Yaskawa INFORM job: OVERLAP3.JBI

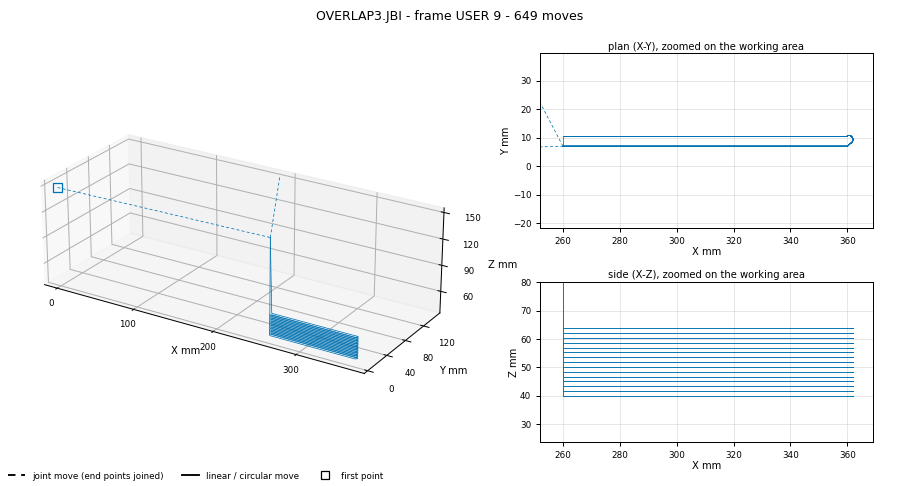
[picture p0: tool path of OVERLAP3.JBI in frame USER 9, 649 of 664 moves have a stored position in this frame; points joined in program order, loops and branches not executed]
/JOB
//NAME OVERLAP1
//POS
///NPOS 664,0,0,0,0,0
///USER 9
///TOOL 1
///POSTYPE USER
///RECTAN
///RCONF 1,0,0,0,0,0,0,0,0,0,0,0,0,0,0,0,0,0,0,0,0,0,0,0
C00000=0.000,0.000,150.000,0.0000,0.0000,45.0000
C00001=260.000,7.000,150.000,0.0000,0.0000,45.0000
C00002=260.000,7.000,40.000,0.0000,0.0000,45.0000
C00003=265.000,7.000,40.000,0.0000,0.0000,45.0000
C00004=270.000,7.000,40.000,0.0000,0.0000,45.0000
C00005=275.000,7.000,40.000,0.0000,0.0000,45.0000
C00006=280.000,7.000,40.000,0.0000,0.0000,45.0000
C00007=285.000,7.000,40.000,0.0000,0.0000,45.0000
C00008=290.000,7.000,40.000,0.0000,0.0000,45.0000
C00009=295.000,7.000,40.000,0.0000,0.0000,45.0000
C00010=300.000,7.000,40.000,0.0000,0.0000,45.0000
C00011=305.000,7.000,40.000,0.0000,0.0000,45.0000
C00012=310.000,7.000,40.000,0.0000,0.0000,45.0000
C00013=315.000,7.000,40.000,0.0000,0.0000,45.0000
C00014=320.000,7.000,40.000,0.0000,0.0000,45.0000
C00015=325.000,7.000,40.000,0.0000,0.0000,45.0000
C00016=330.000,7.000,40.000,0.0000,0.0000,45.0000
C00017=335.000,7.000,40.000,0.0000,0.0000,45.0000
C00018=340.000,7.000,40.000,0.0000,0.0000,45.0000
C00019=345.000,7.000,40.000,0.0000,0.0000,45.0000
C00020=350.000,7.000,40.000,0.0000,0.0000,45.0000
C00021=355.000,7.000,40.000,0.0000,0.0000,45.0000
C00022=360.000,7.000,40.000,0.0000,0.0000,45.0000
C00023=360.938,7.938,40.000,0.0000,0.0000,45.0000
C00024=361.875,9.812,40.000,0.0000,0.0000,45.0000
C00025=360.000,10.750,40.000,0.0000,0.0000,45.0000
C00026=355.000,10.750,40.000,0.0000,0.0000,45.0000
C00027=350.000,10.750,40.000,0.0000,0.0000,45.0000
C00028=345.000,10.750,40.000,0.0000,0.0000,45.0000
C00029=340.000,10.750,40.000,0.0000,0.0000,45.0000
C00030=335.000,10.750,40.000,0.0000,0.0000,45.0000
C00031=330.000,10.750,40.000,0.0000,0.0000,45.0000
C00032=325.000,10.750,40.000,0.0000,0.0000,45.0000
C00033=320.000,10.750,40.000,0.0000,0.0000,45.0000
C00034=315.000,10.750,40.000,0.0000,0.0000,45.0000
C00035=310.000,10.750,40.000,0.0000,0.0000,45.0000
C00036=305.000,10.750,40.000,0.0000,0.0000,45.0000
C00037=300.000,10.750,40.000,0.0000,0.0000,45.0000
C00038=295.000,10.750,40.000,0.0000,0.0000,45.0000
C00039=290.000,10.750,40.000,0.0000,0.0000,45.0000
C00040=285.000,10.750,40.000,0.0000,0.0000,45.0000
C00041=280.000,10.750,40.000,0.0000,0.0000,45.0000
C00042=275.000,10.750,40.000,0.0000,0.0000,45.0000
C00043=270.000,10.750,40.000,0.0000,0.0000,45.0000
C00044=265.000,10.750,40.000,0.0000,0.0000,45.0000
C00045=260.000,10.750,40.000,0.0000,0.0000,45.0000
C00046=260.000,10.750,41.700,0.0000,0.0000,45.0000
C00047=265.000,10.750,41.700,0.0000,0.0000,45.0000
C00048=270.000,10.750,41.700,0.0000,0.0000,45.0000
C00049=275.000,10.750,41.700,0.0000,0.0000,45.0000
C00050=280.000,10.750,41.700,0.0000,0.0000,45.0000
C00051=285.000,10.750,41.700,0.0000,0.0000,45.0000
C00052=290.000,10.750,41.700,0.0000,0.0000,45.0000
C00053=295.000,10.750,41.700,0.0000,0.0000,45.0000
C00054=300.000,10.750,41.700,0.0000,0.0000,45.0000
C00055=305.000,10.750,41.700,0.0000,0.0000,45.0000
C00056=310.000,10.750,41.700,0.0000,0.0000,45.0000
C00057=315.000,10.750,41.700,0.0000,0.0000,45.0000
C00058=320.000,10.750,41.700,0.0000,0.0000,45.0000
C00059=325.000,10.750,41.700,0.0000,0.0000,45.0000
C00060=330.000,10.750,41.700,0.0000,0.0000,45.0000
C00061=335.000,10.750,41.700,0.0000,0.0000,45.0000
C00062=340.000,10.750,41.700,0.0000,0.0000,45.0000
C00063=345.000,10.750,41.700,0.0000,0.0000,45.0000
C00064=350.000,10.750,41.700,0.0000,0.0000,45.0000
C00065=355.000,10.750,41.700,0.0000,0.0000,45.0000
C00066=360.000,10.750,41.700,0.0000,0.0000,45.0000
C00067=361.875,9.812,41.700,0.0000,0.0000,45.0000
C00068=360.938,7.938,41.700,0.0000,0.0000,45.0000
C00069=360.000,7.000,41.700,0.0000,0.0000,45.0000
C00070=355.000,7.000,41.700,0.0000,0.0000,45.0000
C00071=350.000,7.000,41.700,0.0000,0.0000,45.0000
C00072=345.000,7.000,41.700,0.0000,0.0000,45.0000
C00073=340.000,7.000,41.700,0.0000,0.0000,45.0000
C00074=335.000,7.000,41.700,0.0000,0.0000,45.0000
C00075=330.000,7.000,41.700,0.0000,0.0000,45.0000
C00076=325.000,7.000,41.700,0.0000,0.0000,45.0000
C00077=320.000,7.000,41.700,0.0000,0.0000,45.0000
C00078=315.000,7.000,41.700,0.0000,0.0000,45.0000
C00079=310.000,7.000,41.700,0.0000,0.0000,45.0000
C00080=305.000,7.000,41.700,0.0000,0.0000,45.0000
C00081=300.000,7.000,41.700,0.0000,0.0000,45.0000
C00082=295.000,7.000,41.700,0.0000,0.0000,45.0000
C00083=290.000,7.000,41.700,0.0000,0.0000,45.0000
C00084=285.000,7.000,41.700,0.0000,0.0000,45.0000
C00085=280.000,7.000,41.700,0.0000,0.0000,45.0000
C00086=275.000,7.000,41.700,0.0000,0.0000,45.0000
C00087=270.000,7.000,41.700,0.0000,0.0000,45.0000
C00088=265.000,7.000,41.700,0.0000,0.0000,45.0000
C00089=260.000,7.000,41.700,0.0000,0.0000,45.0000
C00090=260.000,7.000,43.400,0.0000,0.0000,45.0000
C00091=265.000,7.000,43.400,0.0000,0.0000,45.0000
C00092=270.000,7.000,43.400,0.0000,0.0000,45.0000
C00093=275.000,7.000,43.400,0.0000,0.0000,45.0000
C00094=280.000,7.000,43.400,0.0000,0.0000,45.0000
C00095=285.000,7.000,43.400,0.0000,0.0000,45.0000
C00096=290.000,7.000,43.400,0.0000,0.0000,45.0000
C00097=295.000,7.000,43.400,0.0000,0.0000,45.0000
C00098=300.000,7.000,43.400,0.0000,0.0000,45.0000
C00099=305.000,7.000,43.400,0.0000,0.0000,45.0000
C00100=310.000,7.000,43.400,0.0000,0.0000,45.0000
C00101=315.000,7.000,43.400,0.0000,0.0000,45.0000
C00102=320.000,7.000,43.400,0.0000,0.0000,45.0000
C00103=325.000,7.000,43.400,0.0000,0.0000,45.0000
C00104=330.000,7.000,43.400,0.0000,0.0000,45.0000
C00105=335.000,7.000,43.400,0.0000,0.0000,45.0000
C00106=340.000,7.000,43.400,0.0000,0.0000,45.0000
C00107=345.000,7.000,43.400,0.0000,0.0000,45.0000
C00108=350.000,7.000,43.400,0.0000,0.0000,45.0000
C00109=355.000,7.000,43.400,0.0000,0.0000,45.0000
C00110=360.000,7.000,43.400,0.0000,0.0000,45.0000
C00111=360.938,7.938,43.400,0.0000,0.0000,45.0000
C00112=361.875,9.812,43.400,0.0000,0.0000,45.0000
C00113=360.000,10.750,43.400,0.0000,0.0000,45.0000
C00114=355.000,10.750,43.400,0.0000,0.0000,45.0000
C00115=350.000,10.750,43.400,0.0000,0.0000,45.0000
C00116=345.000,10.750,43.400,0.0000,0.0000,45.0000
C00117=340.000,10.750,43.400,0.0000,0.0000,45.0000
C00118=335.000,10.750,43.400,0.0000,0.0000,45.0000
C00119=330.000,10.750,43.400,0.0000,0.0000,45.0000
C00120=325.000,10.750,43.400,0.0000,0.0000,45.0000
C00121=320.000,10.750,43.400,0.0000,0.0000,45.0000
C00122=315.000,10.750,43.400,0.0000,0.0000,45.0000
C00123=310.000,10.750,43.400,0.0000,0.0000,45.0000
C00124=305.000,10.750,43.400,0.0000,0.0000,45.0000
C00125=300.000,10.750,43.400,0.0000,0.0000,45.0000
C00126=295.000,10.750,43.400,0.0000,0.0000,45.0000
C00127=290.000,10.750,43.400,0.0000,0.0000,45.0000
C00128=285.000,10.750,43.400,0.0000,0.0000,45.0000
C00129=280.000,10.750,43.400,0.0000,0.0000,45.0000
C00130=275.000,10.750,43.400,0.0000,0.0000,45.0000
C00131=270.000,10.750,43.400,0.0000,0.0000,45.0000
C00132=265.000,10.750,43.400,0.0000,0.0000,45.0000
C00133=260.000,10.750,43.400,0.0000,0.0000,45.0000
C00134=260.000,10.750,45.100,0.0000,0.0000,45.0000
C00135=265.000,10.750,45.100,0.0000,0.0000,45.0000
C00136=270.000,10.750,45.100,0.0000,0.0000,45.0000
C00137=275.000,10.750,45.100,0.0000,0.0000,45.0000
C00138=280.000,10.750,45.100,0.0000,0.0000,45.0000
C00139=285.000,10.750,45.100,0.0000,0.0000,45.0000
C00140=290.000,10.750,45.100,0.0000,0.0000,45.0000
C00141=295.000,10.750,45.100,0.0000,0.0000,45.0000
C00142=300.000,10.750,45.100,0.0000,0.0000,45.0000
C00143=305.000,10.750,45.100,0.0000,0.0000,45.0000
C00144=310.000,10.750,45.100,0.0000,0.0000,45.0000
C00145=315.000,10.750,45.100,0.0000,0.0000,45.0000
C00146=320.000,10.750,45.100,0.0000,0.0000,45.0000
C00147=325.000,10.750,45.100,0.0000,0.0000,45.0000
C00148=330.000,10.750,45.100,0.0000,0.0000,45.0000
C00149=335.000,10.750,45.100,0.0000,0.0000,45.0000
C00150=340.000,10.750,45.100,0.0000,0.0000,45.0000
C00151=345.000,10.750,45.100,0.0000,0.0000,45.0000
C00152=350.000,10.750,45.100,0.0000,0.0000,45.0000
C00153=355.000,10.750,45.100,0.0000,0.0000,45.0000
C00154=360.000,10.750,45.100,0.0000,0.0000,45.0000
C00155=361.875,9.812,45.100,0.0000,0.0000,45.0000
C00156=360.938,7.938,45.100,0.0000,0.0000,45.0000
C00157=360.000,7.000,45.100,0.0000,0.0000,45.0000
C00158=355.000,7.000,45.100,0.0000,0.0000,45.0000
C00159=350.000,7.000,45.100,0.0000,0.0000,45.0000
C00160=345.000,7.000,45.100,0.0000,0.0000,45.0000
C00161=340.000,7.000,45.100,0.0000,0.0000,45.0000
C00162=335.000,7.000,45.100,0.0000,0.0000,45.0000
C00163=330.000,7.000,45.100,0.0000,0.0000,45.0000
C00164=325.000,7.000,45.100,0.0000,0.0000,45.0000
C00165=320.000,7.000,45.100,0.0000,0.0000,45.0000
C00166=315.000,7.000,45.100,0.0000,0.0000,45.0000
C00167=310.000,7.000,45.100,0.0000,0.0000,45.0000
C00168=305.000,7.000,45.100,0.0000,0.0000,45.0000
C00169=300.000,7.000,45.100,0.0000,0.0000,45.0000
C00170=295.000,7.000,45.100,0.0000,0.0000,45.0000
C00171=290.000,7.000,45.100,0.0000,0.0000,45.0000
C00172=285.000,7.000,45.100,0.0000,0.0000,45.0000
C00173=280.000,7.000,45.100,0.0000,0.0000,45.0000
C00174=275.000,7.000,45.100,0.0000,0.0000,45.0000
C00175=270.000,7.000,45.100,0.0000,0.0000,45.0000
C00176=265.000,7.000,45.100,0.0000,0.0000,45.0000
C00177=260.000,7.000,45.100,0.0000,0.0000,45.0000
C00178=260.000,7.000,46.800,0.0000,0.0000,45.0000
C00179=265.000,7.000,46.800,0.0000,0.0000,45.0000
C00180=270.000,7.000,46.800,0.0000,0.0000,45.0000
C00181=275.000,7.000,46.800,0.0000,0.0000,45.0000
C00182=280.000,7.000,46.800,0.0000,0.0000,45.0000
C00183=285.000,7.000,46.800,0.0000,0.0000,45.0000
C00184=290.000,7.000,46.800,0.0000,0.0000,45.0000
C00185=295.000,7.000,46.800,0.0000,0.0000,45.0000
C00186=300.000,7.000,46.800,0.0000,0.0000,45.0000
C00187=305.000,7.000,46.800,0.0000,0.0000,45.0000
C00188=310.000,7.000,46.800,0.0000,0.0000,45.0000
C00189=315.000,7.000,46.800,0.0000,0.0000,45.0000
C00190=320.000,7.000,46.800,0.0000,0.0000,45.0000
C00191=325.000,7.000,46.800,0.0000,0.0000,45.0000
C00192=330.000,7.000,46.800,0.0000,0.0000,45.0000
C00193=335.000,7.000,46.800,0.0000,0.0000,45.0000
C00194=340.000,7.000,46.800,0.0000,0.0000,45.0000
C00195=345.000,7.000,46.800,0.0000,0.0000,45.0000
C00196=350.000,7.000,46.800,0.0000,0.0000,45.0000
C00197=355.000,7.000,46.800,0.0000,0.0000,45.0000
C00198=360.000,7.000,46.800,0.0000,0.0000,45.0000
C00199=360.938,7.938,46.800,0.0000,0.0000,45.0000
C00200=361.875,9.812,46.800,0.0000,0.0000,45.0000
C00201=360.000,10.750,46.800,0.0000,0.0000,45.0000
C00202=355.000,10.750,46.800,0.0000,0.0000,45.0000
C00203=350.000,10.750,46.800,0.0000,0.0000,45.0000
C00204=345.000,10.750,46.800,0.0000,0.0000,45.0000
C00205=340.000,10.750,46.800,0.0000,0.0000,45.0000
C00206=335.000,10.750,46.800,0.0000,0.0000,45.0000
C00207=330.000,10.750,46.800,0.0000,0.0000,45.0000
C00208=325.000,10.750,46.800,0.0000,0.0000,45.0000
C00209=320.000,10.750,46.800,0.0000,0.0000,45.0000
C00210=315.000,10.750,46.800,0.0000,0.0000,45.0000
C00211=310.000,10.750,46.800,0.0000,0.0000,45.0000
C00212=305.000,10.750,46.800,0.0000,0.0000,45.0000
C00213=300.000,10.750,46.800,0.0000,0.0000,45.0000
C00214=295.000,10.750,46.800,0.0000,0.0000,45.0000
C00215=290.000,10.750,46.800,0.0000,0.0000,45.0000
C00216=285.000,10.750,46.800,0.0000,0.0000,45.0000
C00217=280.000,10.750,46.800,0.0000,0.0000,45.0000
C00218=275.000,10.750,46.800,0.0000,0.0000,45.0000
C00219=270.000,10.750,46.800,0.0000,0.0000,45.0000
C00220=265.000,10.750,46.800,0.0000,0.0000,45.0000
C00221=260.000,10.750,46.800,0.0000,0.0000,45.0000
C00222=260.000,10.750,48.500,0.0000,0.0000,45.0000
C00223=265.000,10.750,48.500,0.0000,0.0000,45.0000
C00224=270.000,10.750,48.500,0.0000,0.0000,45.0000
C00225=275.000,10.750,48.500,0.0000,0.0000,45.0000
C00226=280.000,10.750,48.500,0.0000,0.0000,45.0000
C00227=285.000,10.750,48.500,0.0000,0.0000,45.0000
C00228=290.000,10.750,48.500,0.0000,0.0000,45.0000
C00229=295.000,10.750,48.500,0.0000,0.0000,45.0000
C00230=300.000,10.750,48.500,0.0000,0.0000,45.0000
C00231=305.000,10.750,48.500,0.0000,0.0000,45.0000
C00232=310.000,10.750,48.500,0.0000,0.0000,45.0000
C00233=315.000,10.750,48.500,0.0000,0.0000,45.0000
C00234=320.000,10.750,48.500,0.0000,0.0000,45.0000
C00235=325.000,10.750,48.500,0.0000,0.0000,45.0000
C00236=330.000,10.750,48.500,0.0000,0.0000,45.0000
C00237=335.000,10.750,48.500,0.0000,0.0000,45.0000
C00238=340.000,10.750,48.500,0.0000,0.0000,45.0000
C00239=345.000,10.750,48.500,0.0000,0.0000,45.0000
C00240=350.000,10.750,48.500,0.0000,0.0000,45.0000
C00241=355.000,10.750,48.500,0.0000,0.0000,45.0000
C00242=360.000,10.750,48.500,0.0000,0.0000,45.0000
C00243=361.875,9.812,48.500,0.0000,0.0000,45.0000
C00244=360.938,7.938,48.500,0.0000,0.0000,45.0000
C00245=360.000,7.000,48.500,0.0000,0.0000,45.0000
C00246=355.000,7.000,48.500,0.0000,0.0000,45.0000
C00247=350.000,7.000,48.500,0.0000,0.0000,45.0000
C00248=345.000,7.000,48.500,0.0000,0.0000,45.0000
C00249=340.000,7.000,48.500,0.0000,0.0000,45.0000
C00250=335.000,7.000,48.500,0.0000,0.0000,45.0000
C00251=330.000,7.000,48.500,0.0000,0.0000,45.0000
C00252=325.000,7.000,48.500,0.0000,0.0000,45.0000
C00253=320.000,7.000,48.500,0.0000,0.0000,45.0000
C00254=315.000,7.000,48.500,0.0000,0.0000,45.0000
C00255=310.000,7.000,48.500,0.0000,0.0000,45.0000
C00256=305.000,7.000,48.500,0.0000,0.0000,45.0000
C00257=300.000,7.000,48.500,0.0000,0.0000,45.0000
C00258=295.000,7.000,48.500,0.0000,0.0000,45.0000
C00259=290.000,7.000,48.500,0.0000,0.0000,45.0000
C00260=285.000,7.000,48.500,0.0000,0.0000,45.0000
C00261=280.000,7.000,48.500,0.0000,0.0000,45.0000
C00262=275.000,7.000,48.500,0.0000,0.0000,45.0000
C00263=270.000,7.000,48.500,0.0000,0.0000,45.0000
C00264=265.000,7.000,48.500,0.0000,0.0000,45.0000
C00265=260.000,7.000,48.500,0.0000,0.0000,45.0000
C00266=260.000,7.000,50.200,0.0000,0.0000,45.0000
C00267=265.000,7.000,50.200,0.0000,0.0000,45.0000
C00268=270.000,7.000,50.200,0.0000,0.0000,45.0000
C00269=275.000,7.000,50.200,0.0000,0.0000,45.0000
C00270=280.000,7.000,50.200,0.0000,0.0000,45.0000
C00271=285.000,7.000,50.200,0.0000,0.0000,45.0000
C00272=290.000,7.000,50.200,0.0000,0.0000,45.0000
C00273=295.000,7.000,50.200,0.0000,0.0000,45.0000
C00274=300.000,7.000,50.200,0.0000,0.0000,45.0000
C00275=305.000,7.000,50.200,0.0000,0.0000,45.0000
C00276=310.000,7.000,50.200,0.0000,0.0000,45.0000
C00277=315.000,7.000,50.200,0.0000,0.0000,45.0000
C00278=320.000,7.000,50.200,0.0000,0.0000,45.0000
C00279=325.000,7.000,50.200,0.0000,0.0000,45.0000
C00280=330.000,7.000,50.200,0.0000,0.0000,45.0000
C00281=335.000,7.000,50.200,0.0000,0.0000,45.0000
C00282=340.000,7.000,50.200,0.0000,0.0000,45.0000
C00283=345.000,7.000,50.200,0.0000,0.0000,45.0000
C00284=350.000,7.000,50.200,0.0000,0.0000,45.0000
C00285=355.000,7.000,50.200,0.0000,0.0000,45.0000
C00286=360.000,7.000,50.200,0.0000,0.0000,45.0000
C00287=360.938,7.938,50.200,0.0000,0.0000,45.0000
C00288=361.875,9.812,50.200,0.0000,0.0000,45.0000
C00289=360.000,10.750,50.200,0.0000,0.0000,45.0000
C00290=355.000,10.750,50.200,0.0000,0.0000,45.0000
C00291=350.000,10.750,50.200,0.0000,0.0000,45.0000
C00292=345.000,10.750,50.200,0.0000,0.0000,45.0000
C00293=340.000,10.750,50.200,0.0000,0.0000,45.0000
C00294=335.000,10.750,50.200,0.0000,0.0000,45.0000
C00295=330.000,10.750,50.200,0.0000,0.0000,45.0000
C00296=325.000,10.750,50.200,0.0000,0.0000,45.0000
C00297=320.000,10.750,50.200,0.0000,0.0000,45.0000
C00298=315.000,10.750,50.200,0.0000,0.0000,45.0000
C00299=310.000,10.750,50.200,0.0000,0.0000,45.0000
C00300=305.000,10.750,50.200,0.0000,0.0000,45.0000
C00301=300.000,10.750,50.200,0.0000,0.0000,45.0000
C00302=295.000,10.750,50.200,0.0000,0.0000,45.0000
C00303=290.000,10.750,50.200,0.0000,0.0000,45.0000
C00304=285.000,10.750,50.200,0.0000,0.0000,45.0000
C00305=280.000,10.750,50.200,0.0000,0.0000,45.0000
C00306=275.000,10.750,50.200,0.0000,0.0000,45.0000
C00307=270.000,10.750,50.200,0.0000,0.0000,45.0000
C00308=265.000,10.750,50.200,0.0000,0.0000,45.0000
C00309=260.000,10.750,50.200,0.0000,0.0000,45.0000
C00310=260.000,10.750,51.900,0.0000,0.0000,45.0000
C00311=265.000,10.750,51.900,0.0000,0.0000,45.0000
C00312=270.000,10.750,51.900,0.0000,0.0000,45.0000
C00313=275.000,10.750,51.900,0.0000,0.0000,45.0000
C00314=280.000,10.750,51.900,0.0000,0.0000,45.0000
C00315=285.000,10.750,51.900,0.0000,0.0000,45.0000
C00316=290.000,10.750,51.900,0.0000,0.0000,45.0000
C00317=295.000,10.750,51.900,0.0000,0.0000,45.0000
C00318=300.000,10.750,51.900,0.0000,0.0000,45.0000
C00319=305.000,10.750,51.900,0.0000,0.0000,45.0000
C00320=310.000,10.750,51.900,0.0000,0.0000,45.0000
C00321=315.000,10.750,51.900,0.0000,0.0000,45.0000
C00322=320.000,10.750,51.900,0.0000,0.0000,45.0000
C00323=325.000,10.750,51.900,0.0000,0.0000,45.0000
C00324=330.000,10.750,51.900,0.0000,0.0000,45.0000
C00325=335.000,10.750,51.900,0.0000,0.0000,45.0000
C00326=340.000,10.750,51.900,0.0000,0.0000,45.0000
C00327=345.000,10.750,51.900,0.0000,0.0000,45.0000
C00328=350.000,10.750,51.900,0.0000,0.0000,45.0000
C00329=355.000,10.750,51.900,0.0000,0.0000,45.0000
C00330=360.000,10.750,51.900,0.0000,0.0000,45.0000
C00331=361.875,9.812,51.900,0.0000,0.0000,45.0000
C00332=360.938,7.938,51.900,0.0000,0.0000,45.0000
C00333=360.000,7.000,51.900,0.0000,0.0000,45.0000
C00334=355.000,7.000,51.900,0.0000,0.0000,45.0000
C00335=350.000,7.000,51.900,0.0000,0.0000,45.0000
C00336=345.000,7.000,51.900,0.0000,0.0000,45.0000
C00337=340.000,7.000,51.900,0.0000,0.0000,45.0000
C00338=335.000,7.000,51.900,0.0000,0.0000,45.0000
C00339=330.000,7.000,51.900,0.0000,0.0000,45.0000
C00340=325.000,7.000,51.900,0.0000,0.0000,45.0000
C00341=320.000,7.000,51.900,0.0000,0.0000,45.0000
C00342=315.000,7.000,51.900,0.0000,0.0000,45.0000
C00343=310.000,7.000,51.900,0.0000,0.0000,45.0000
C00344=305.000,7.000,51.900,0.0000,0.0000,45.0000
C00345=300.000,7.000,51.900,0.0000,0.0000,45.0000
C00346=295.000,7.000,51.900,0.0000,0.0000,45.0000
C00347=290.000,7.000,51.900,0.0000,0.0000,45.0000
C00348=285.000,7.000,51.900,0.0000,0.0000,45.0000
C00349=280.000,7.000,51.900,0.0000,0.0000,45.0000
C00350=275.000,7.000,51.900,0.0000,0.0000,45.0000
C00351=270.000,7.000,51.900,0.0000,0.0000,45.0000
C00352=265.000,7.000,51.900,0.0000,0.0000,45.0000
C00353=260.000,7.000,51.900,0.0000,0.0000,45.0000
C00354=260.000,7.000,53.600,0.0000,0.0000,45.0000
C00355=265.000,7.000,53.600,0.0000,0.0000,45.0000
C00356=270.000,7.000,53.600,0.0000,0.0000,45.0000
C00357=275.000,7.000,53.600,0.0000,0.0000,45.0000
C00358=280.000,7.000,53.600,0.0000,0.0000,45.0000
C00359=285.000,7.000,53.600,0.0000,0.0000,45.0000
C00360=290.000,7.000,53.600,0.0000,0.0000,45.0000
C00361=295.000,7.000,53.600,0.0000,0.0000,45.0000
C00362=300.000,7.000,53.600,0.0000,0.0000,45.0000
C00363=305.000,7.000,53.600,0.0000,0.0000,45.0000
C00364=310.000,7.000,53.600,0.0000,0.0000,45.0000
C00365=315.000,7.000,53.600,0.0000,0.0000,45.0000
C00366=320.000,7.000,53.600,0.0000,0.0000,45.0000
C00367=325.000,7.000,53.600,0.0000,0.0000,45.0000
C00368=330.000,7.000,53.600,0.0000,0.0000,45.0000
C00369=335.000,7.000,53.600,0.0000,0.0000,45.0000
C00370=340.000,7.000,53.600,0.0000,0.0000,45.0000
C00371=345.000,7.000,53.600,0.0000,0.0000,45.0000
C00372=350.000,7.000,53.600,0.0000,0.0000,45.0000
C00373=355.000,7.000,53.600,0.0000,0.0000,45.0000
C00374=360.000,7.000,53.600,0.0000,0.0000,45.0000
C00375=360.938,7.938,53.600,0.0000,0.0000,45.0000
C00376=361.875,9.812,53.600,0.0000,0.0000,45.0000
C00377=360.000,10.750,53.600,0.0000,0.0000,45.0000
C00378=355.000,10.750,53.600,0.0000,0.0000,45.0000
C00379=350.000,10.750,53.600,0.0000,0.0000,45.0000
C00380=345.000,10.750,53.600,0.0000,0.0000,45.0000
C00381=340.000,10.750,53.600,0.0000,0.0000,45.0000
C00382=335.000,10.750,53.600,0.0000,0.0000,45.0000
C00383=330.000,10.750,53.600,0.0000,0.0000,45.0000
C00384=325.000,10.750,53.600,0.0000,0.0000,45.0000
C00385=320.000,10.750,53.600,0.0000,0.0000,45.0000
C00386=315.000,10.750,53.600,0.0000,0.0000,45.0000
C00387=310.000,10.750,53.600,0.0000,0.0000,45.0000
C00388=305.000,10.750,53.600,0.0000,0.0000,45.0000
C00389=300.000,10.750,53.600,0.0000,0.0000,45.0000
C00390=295.000,10.750,53.600,0.0000,0.0000,45.0000
C00391=290.000,10.750,53.600,0.0000,0.0000,45.0000
C00392=285.000,10.750,53.600,0.0000,0.0000,45.0000
C00393=280.000,10.750,53.600,0.0000,0.0000,45.0000
C00394=275.000,10.750,53.600,0.0000,0.0000,45.0000
C00395=270.000,10.750,53.600,0.0000,0.0000,45.0000
C00396=265.000,10.750,53.600,0.0000,0.0000,45.0000
C00397=260.000,10.750,53.600,0.0000,0.0000,45.0000
C00398=260.000,10.750,55.300,0.0000,0.0000,45.0000
C00399=265.000,10.750,55.300,0.0000,0.0000,45.0000
C00400=270.000,10.750,55.300,0.0000,0.0000,45.0000
C00401=275.000,10.750,55.300,0.0000,0.0000,45.0000
C00402=280.000,10.750,55.300,0.0000,0.0000,45.0000
C00403=285.000,10.750,55.300,0.0000,0.0000,45.0000
C00404=290.000,10.750,55.300,0.0000,0.0000,45.0000
C00405=295.000,10.750,55.300,0.0000,0.0000,45.0000
C00406=300.000,10.750,55.300,0.0000,0.0000,45.0000
C00407=305.000,10.750,55.300,0.0000,0.0000,45.0000
C00408=310.000,10.750,55.300,0.0000,0.0000,45.0000
C00409=315.000,10.750,55.300,0.0000,0.0000,45.0000
C00410=320.000,10.750,55.300,0.0000,0.0000,45.0000
C00411=325.000,10.750,55.300,0.0000,0.0000,45.0000
C00412=330.000,10.750,55.300,0.0000,0.0000,45.0000
C00413=335.000,10.750,55.300,0.0000,0.0000,45.0000
C00414=340.000,10.750,55.300,0.0000,0.0000,45.0000
C00415=345.000,10.750,55.300,0.0000,0.0000,45.0000
C00416=350.000,10.750,55.300,0.0000,0.0000,45.0000
C00417=355.000,10.750,55.300,0.0000,0.0000,45.0000
C00418=360.000,10.750,55.300,0.0000,0.0000,45.0000
C00419=361.875,9.812,55.300,0.0000,0.0000,45.0000
C00420=360.938,7.938,55.300,0.0000,0.0000,45.0000
C00421=360.000,7.000,55.300,0.0000,0.0000,45.0000
C00422=355.000,7.000,55.300,0.0000,0.0000,45.0000
C00423=350.000,7.000,55.300,0.0000,0.0000,45.0000
C00424=345.000,7.000,55.300,0.0000,0.0000,45.0000
C00425=340.000,7.000,55.300,0.0000,0.0000,45.0000
C00426=335.000,7.000,55.300,0.0000,0.0000,45.0000
C00427=330.000,7.000,55.300,0.0000,0.0000,45.0000
C00428=325.000,7.000,55.300,0.0000,0.0000,45.0000
C00429=320.000,7.000,55.300,0.0000,0.0000,45.0000
C00430=315.000,7.000,55.300,0.0000,0.0000,45.0000
C00431=310.000,7.000,55.300,0.0000,0.0000,45.0000
C00432=305.000,7.000,55.300,0.0000,0.0000,45.0000
C00433=300.000,7.000,55.300,0.0000,0.0000,45.0000
C00434=295.000,7.000,55.300,0.0000,0.0000,45.0000
C00435=290.000,7.000,55.300,0.0000,0.0000,45.0000
C00436=285.000,7.000,55.300,0.0000,0.0000,45.0000
C00437=280.000,7.000,55.300,0.0000,0.0000,45.0000
C00438=275.000,7.000,55.300,0.0000,0.0000,45.0000
C00439=270.000,7.000,55.300,0.0000,0.0000,45.0000
C00440=265.000,7.000,55.300,0.0000,0.0000,45.0000
C00441=260.000,7.000,55.300,0.0000,0.0000,45.0000
C00442=260.000,7.000,57.000,0.0000,0.0000,45.0000
C00443=265.000,7.000,57.000,0.0000,0.0000,45.0000
C00444=270.000,7.000,57.000,0.0000,0.0000,45.0000
C00445=275.000,7.000,57.000,0.0000,0.0000,45.0000
C00446=280.000,7.000,57.000,0.0000,0.0000,45.0000
C00447=285.000,7.000,57.000,0.0000,0.0000,45.0000
C00448=290.000,7.000,57.000,0.0000,0.0000,45.0000
C00449=295.000,7.000,57.000,0.0000,0.0000,45.0000
C00450=300.000,7.000,57.000,0.0000,0.0000,45.0000
C00451=305.000,7.000,57.000,0.0000,0.0000,45.0000
C00452=310.000,7.000,57.000,0.0000,0.0000,45.0000
C00453=315.000,7.000,57.000,0.0000,0.0000,45.0000
C00454=320.000,7.000,57.000,0.0000,0.0000,45.0000
C00455=325.000,7.000,57.000,0.0000,0.0000,45.0000
C00456=330.000,7.000,57.000,0.0000,0.0000,45.0000
C00457=335.000,7.000,57.000,0.0000,0.0000,45.0000
C00458=340.000,7.000,57.000,0.0000,0.0000,45.0000
C00459=345.000,7.000,57.000,0.0000,0.0000,45.0000
C00460=350.000,7.000,57.000,0.0000,0.0000,45.0000
C00461=355.000,7.000,57.000,0.0000,0.0000,45.0000
C00462=360.000,7.000,57.000,0.0000,0.0000,45.0000
C00463=360.938,7.938,57.000,0.0000,0.0000,45.0000
C00464=361.875,9.812,57.000,0.0000,0.0000,45.0000
C00465=360.000,10.750,57.000,0.0000,0.0000,45.0000
C00466=355.000,10.750,57.000,0.0000,0.0000,45.0000
C00467=350.000,10.750,57.000,0.0000,0.0000,45.0000
C00468=345.000,10.750,57.000,0.0000,0.0000,45.0000
C00469=340.000,10.750,57.000,0.0000,0.0000,45.0000
C00470=335.000,10.750,57.000,0.0000,0.0000,45.0000
C00471=330.000,10.750,57.000,0.0000,0.0000,45.0000
C00472=325.000,10.750,57.000,0.0000,0.0000,45.0000
C00473=320.000,10.750,57.000,0.0000,0.0000,45.0000
C00474=315.000,10.750,57.000,0.0000,0.0000,45.0000
C00475=310.000,10.750,57.000,0.0000,0.0000,45.0000
C00476=305.000,10.750,57.000,0.0000,0.0000,45.0000
C00477=300.000,10.750,57.000,0.0000,0.0000,45.0000
C00478=295.000,10.750,57.000,0.0000,0.0000,45.0000
C00479=290.000,10.750,57.000,0.0000,0.0000,45.0000
C00480=285.000,10.750,57.000,0.0000,0.0000,45.0000
C00481=280.000,10.750,57.000,0.0000,0.0000,45.0000
C00482=275.000,10.750,57.000,0.0000,0.0000,45.0000
C00483=270.000,10.750,57.000,0.0000,0.0000,45.0000
C00484=265.000,10.750,57.000,0.0000,0.0000,45.0000
C00485=260.000,10.750,57.000,0.0000,0.0000,45.0000
C00486=260.000,10.750,58.700,0.0000,0.0000,45.0000
C00487=265.000,10.750,58.700,0.0000,0.0000,45.0000
C00488=270.000,10.750,58.700,0.0000,0.0000,45.0000
C00489=275.000,10.750,58.700,0.0000,0.0000,45.0000
C00490=280.000,10.750,58.700,0.0000,0.0000,45.0000
C00491=285.000,10.750,58.700,0.0000,0.0000,45.0000
C00492=290.000,10.750,58.700,0.0000,0.0000,45.0000
C00493=295.000,10.750,58.700,0.0000,0.0000,45.0000
C00494=300.000,10.750,58.700,0.0000,0.0000,45.0000
C00495=305.000,10.750,58.700,0.0000,0.0000,45.0000
C00496=310.000,10.750,58.700,0.0000,0.0000,45.0000
C00497=315.000,10.750,58.700,0.0000,0.0000,45.0000
C00498=320.000,10.750,58.700,0.0000,0.0000,45.0000
C00499=325.000,10.750,58.700,0.0000,0.0000,45.0000
C00500=330.000,10.750,58.700,0.0000,0.0000,45.0000
C00501=335.000,10.750,58.700,0.0000,0.0000,45.0000
C00502=340.000,10.750,58.700,0.0000,0.0000,45.0000
C00503=345.000,10.750,58.700,0.0000,0.0000,45.0000
C00504=350.000,10.750,58.700,0.0000,0.0000,45.0000
C00505=355.000,10.750,58.700,0.0000,0.0000,45.0000
C00506=360.000,10.750,58.700,0.0000,0.0000,45.0000
C00507=361.875,9.812,58.700,0.0000,0.0000,45.0000
C00508=360.938,7.938,58.700,0.0000,0.0000,45.0000
C00509=360.000,7.000,58.700,0.0000,0.0000,45.0000
C00510=355.000,7.000,58.700,0.0000,0.0000,45.0000
C00511=350.000,7.000,58.700,0.0000,0.0000,45.0000
C00512=345.000,7.000,58.700,0.0000,0.0000,45.0000
C00513=340.000,7.000,58.700,0.0000,0.0000,45.0000
C00514=335.000,7.000,58.700,0.0000,0.0000,45.0000
C00515=330.000,7.000,58.700,0.0000,0.0000,45.0000
C00516=325.000,7.000,58.700,0.0000,0.0000,45.0000
C00517=320.000,7.000,58.700,0.0000,0.0000,45.0000
C00518=315.000,7.000,58.700,0.0000,0.0000,45.0000
C00519=310.000,7.000,58.700,0.0000,0.0000,45.0000
C00520=305.000,7.000,58.700,0.0000,0.0000,45.0000
C00521=300.000,7.000,58.700,0.0000,0.0000,45.0000
C00522=295.000,7.000,58.700,0.0000,0.0000,45.0000
C00523=290.000,7.000,58.700,0.0000,0.0000,45.0000
C00524=285.000,7.000,58.700,0.0000,0.0000,45.0000
C00525=280.000,7.000,58.700,0.0000,0.0000,45.0000
C00526=275.000,7.000,58.700,0.0000,0.0000,45.0000
C00527=270.000,7.000,58.700,0.0000,0.0000,45.0000
C00528=265.000,7.000,58.700,0.0000,0.0000,45.0000
C00529=260.000,7.000,58.700,0.0000,0.0000,45.0000
C00530=260.000,7.000,60.400,0.0000,0.0000,45.0000
C00531=265.000,7.000,60.400,0.0000,0.0000,45.0000
C00532=270.000,7.000,60.400,0.0000,0.0000,45.0000
C00533=275.000,7.000,60.400,0.0000,0.0000,45.0000
C00534=280.000,7.000,60.400,0.0000,0.0000,45.0000
C00535=285.000,7.000,60.400,0.0000,0.0000,45.0000
C00536=290.000,7.000,60.400,0.0000,0.0000,45.0000
C00537=295.000,7.000,60.400,0.0000,0.0000,45.0000
C00538=300.000,7.000,60.400,0.0000,0.0000,45.0000
C00539=305.000,7.000,60.400,0.0000,0.0000,45.0000
C00540=310.000,7.000,60.400,0.0000,0.0000,45.0000
C00541=315.000,7.000,60.400,0.0000,0.0000,45.0000
C00542=320.000,7.000,60.400,0.0000,0.0000,45.0000
C00543=325.000,7.000,60.400,0.0000,0.0000,45.0000
C00544=330.000,7.000,60.400,0.0000,0.0000,45.0000
C00545=335.000,7.000,60.400,0.0000,0.0000,45.0000
C00546=340.000,7.000,60.400,0.0000,0.0000,45.0000
C00547=345.000,7.000,60.400,0.0000,0.0000,45.0000
C00548=350.000,7.000,60.400,0.0000,0.0000,45.0000
C00549=355.000,7.000,60.400,0.0000,0.0000,45.0000
C00550=360.000,7.000,60.400,0.0000,0.0000,45.0000
C00551=360.938,7.938,60.400,0.0000,0.0000,45.0000
C00552=361.875,9.812,60.400,0.0000,0.0000,45.0000
C00553=360.000,10.750,60.400,0.0000,0.0000,45.0000
C00554=355.000,10.750,60.400,0.0000,0.0000,45.0000
C00555=350.000,10.750,60.400,0.0000,0.0000,45.0000
C00556=345.000,10.750,60.400,0.0000,0.0000,45.0000
C00557=340.000,10.750,60.400,0.0000,0.0000,45.0000
C00558=335.000,10.750,60.400,0.0000,0.0000,45.0000
C00559=330.000,10.750,60.400,0.0000,0.0000,45.0000
C00560=325.000,10.750,60.400,0.0000,0.0000,45.0000
C00561=320.000,10.750,60.400,0.0000,0.0000,45.0000
C00562=315.000,10.750,60.400,0.0000,0.0000,45.0000
C00563=310.000,10.750,60.400,0.0000,0.0000,45.0000
C00564=305.000,10.750,60.400,0.0000,0.0000,45.0000
C00565=300.000,10.750,60.400,0.0000,0.0000,45.0000
C00566=295.000,10.750,60.400,0.0000,0.0000,45.0000
C00567=290.000,10.750,60.400,0.0000,0.0000,45.0000
C00568=285.000,10.750,60.400,0.0000,0.0000,45.0000
C00569=280.000,10.750,60.400,0.0000,0.0000,45.0000
C00570=275.000,10.750,60.400,0.0000,0.0000,45.0000
C00571=270.000,10.750,60.400,0.0000,0.0000,45.0000
C00572=265.000,10.750,60.400,0.0000,0.0000,45.0000
C00573=260.000,10.750,60.400,0.0000,0.0000,45.0000
C00574=260.000,10.750,62.100,0.0000,0.0000,45.0000
C00575=265.000,10.750,62.100,0.0000,0.0000,45.0000
C00576=270.000,10.750,62.100,0.0000,0.0000,45.0000
C00577=275.000,10.750,62.100,0.0000,0.0000,45.0000
C00578=280.000,10.750,62.100,0.0000,0.0000,45.0000
C00579=285.000,10.750,62.100,0.0000,0.0000,45.0000
C00580=290.000,10.750,62.100,0.0000,0.0000,45.0000
C00581=295.000,10.750,62.100,0.0000,0.0000,45.0000
C00582=300.000,10.750,62.100,0.0000,0.0000,45.0000
C00583=305.000,10.750,62.100,0.0000,0.0000,45.0000
C00584=310.000,10.750,62.100,0.0000,0.0000,45.0000
C00585=315.000,10.750,62.100,0.0000,0.0000,45.0000
C00586=320.000,10.750,62.100,0.0000,0.0000,45.0000
C00587=325.000,10.750,62.100,0.0000,0.0000,45.0000
C00588=330.000,10.750,62.100,0.0000,0.0000,45.0000
C00589=335.000,10.750,62.100,0.0000,0.0000,45.0000
C00590=340.000,10.750,62.100,0.0000,0.0000,45.0000
C00591=345.000,10.750,62.100,0.0000,0.0000,45.0000
C00592=350.000,10.750,62.100,0.0000,0.0000,45.0000
C00593=355.000,10.750,62.100,0.0000,0.0000,45.0000
C00594=360.000,10.750,62.100,0.0000,0.0000,45.0000
C00595=361.875,9.812,62.100,0.0000,0.0000,45.0000
C00596=360.938,7.938,62.100,0.0000,0.0000,45.0000
C00597=360.000,7.000,62.100,0.0000,0.0000,45.0000
C00598=355.000,7.000,62.100,0.0000,0.0000,45.0000
C00599=350.000,7.000,62.100,0.0000,0.0000,45.0000
C00600=345.000,7.000,62.100,0.0000,0.0000,45.0000
C00601=340.000,7.000,62.100,0.0000,0.0000,45.0000
C00602=335.000,7.000,62.100,0.0000,0.0000,45.0000
C00603=330.000,7.000,62.100,0.0000,0.0000,45.0000
C00604=325.000,7.000,62.100,0.0000,0.0000,45.0000
C00605=320.000,7.000,62.100,0.0000,0.0000,45.0000
C00606=315.000,7.000,62.100,0.0000,0.0000,45.0000
C00607=310.000,7.000,62.100,0.0000,0.0000,45.0000
C00608=305.000,7.000,62.100,0.0000,0.0000,45.0000
C00609=300.000,7.000,62.100,0.0000,0.0000,45.0000
C00610=295.000,7.000,62.100,0.0000,0.0000,45.0000
C00611=290.000,7.000,62.100,0.0000,0.0000,45.0000
C00612=285.000,7.000,62.100,0.0000,0.0000,45.0000
C00613=280.000,7.000,62.100,0.0000,0.0000,45.0000
C00614=275.000,7.000,62.100,0.0000,0.0000,45.0000
C00615=270.000,7.000,62.100,0.0000,0.0000,45.0000
C00616=265.000,7.000,62.100,0.0000,0.0000,45.0000
C00617=260.000,7.000,62.100,0.0000,0.0000,45.0000
C00618=260.000,7.000,63.800,0.0000,0.0000,45.0000
C00619=265.000,7.000,63.800,0.0000,0.0000,45.0000
C00620=270.000,7.000,63.800,0.0000,0.0000,45.0000
C00621=275.000,7.000,63.800,0.0000,0.0000,45.0000
C00622=280.000,7.000,63.800,0.0000,0.0000,45.0000
C00623=285.000,7.000,63.800,0.0000,0.0000,45.0000
C00624=290.000,7.000,63.800,0.0000,0.0000,45.0000
C00625=295.000,7.000,63.800,0.0000,0.0000,45.0000
C00626=300.000,7.000,63.800,0.0000,0.0000,45.0000
C00627=305.000,7.000,63.800,0.0000,0.0000,45.0000
C00628=310.000,7.000,63.800,0.0000,0.0000,45.0000
C00629=315.000,7.000,63.800,0.0000,0.0000,45.0000
C00630=320.000,7.000,63.800,0.0000,0.0000,45.0000
C00631=325.000,7.000,63.800,0.0000,0.0000,45.0000
C00632=330.000,7.000,63.800,0.0000,0.0000,45.0000
C00633=335.000,7.000,63.800,0.0000,0.0000,45.0000
C00634=340.000,7.000,63.800,0.0000,0.0000,45.0000
C00635=345.000,7.000,63.800,0.0000,0.0000,45.0000
C00636=350.000,7.000,63.800,0.0000,0.0000,45.0000
C00637=355.000,7.000,63.800,0.0000,0.0000,45.0000
C00638=360.000,7.000,63.800,0.0000,0.0000,45.0000
C00639=360.938,7.938,63.800,0.0000,0.0000,45.0000
C00640=361.875,9.812,63.800,0.0000,0.0000,45.0000
C00641=360.000,10.750,63.800,0.0000,0.0000,45.0000
C00642=355.000,10.750,63.800,0.0000,0.0000,45.0000
C00643=350.000,10.750,63.800,0.0000,0.0000,45.0000
C00644=345.000,10.750,63.800,0.0000,0.0000,45.0000
C00645=340.000,10.750,63.800,0.0000,0.0000,45.0000
C00646=335.000,10.750,63.800,0.0000,0.0000,45.0000
C00647=330.000,10.750,63.800,0.0000,0.0000,45.0000
C00648=325.000,10.750,63.800,0.0000,0.0000,45.0000
C00649=320.000,10.750,63.800,0.0000,0.0000,45.0000
C00650=315.000,10.750,63.800,0.0000,0.0000,45.0000
C00651=310.000,10.750,63.800,0.0000,0.0000,45.0000
C00652=305.000,10.750,63.800,0.0000,0.0000,45.0000
C00653=300.000,10.750,63.800,0.0000,0.0000,45.0000
C00654=295.000,10.750,63.800,0.0000,0.0000,45.0000
C00655=290.000,10.750,63.800,0.0000,0.0000,45.0000
C00656=285.000,10.750,63.800,0.0000,0.0000,45.0000
C00657=280.000,10.750,63.800,0.0000,0.0000,45.0000
C00658=275.000,10.750,63.800,0.0000,0.0000,45.0000
C00659=270.000,10.750,63.800,0.0000,0.0000,45.0000
C00660=265.000,10.750,63.800,0.0000,0.0000,45.0000
C00661=260.000,10.750,63.800,0.0000,0.0000,45.0000
C00662=260.000,7.000,150.000,0.0000,0.0000,45.0000
C00663=185.000,150.000,150.000,0.0000,0.0000,45.0000
//INST
///DATE 2026/11/10 11:37
///ATTR SC,RW,RJ
////FRAME USER 9
///GROUP1 RB1
NOP
MOVJ C00000 VJ=0.78
MOVJ C00001 VJ=0.78
MOVL C00002 V=11.0 ACC=20 DEC=20
*LAG1
MACRO1 MJ#(0) ARGF1
ARCON
MOVL C00003 V=7.0 ACC=20 DEC=20
MOVL C00004 V=7.0 ACC=20 DEC=20
MOVL C00005 V=7.0 ACC=20 DEC=20
MOVL C00006 V=7.0 ACC=20 DEC=20
MOVL C00007 V=7.0 ACC=20 DEC=20
MOVL C00008 V=7.0 ACC=20 DEC=20
MOVL C00009 V=7.0 ACC=20 DEC=20
MOVL C00010 V=7.0 ACC=20 DEC=20
MOVL C00011 V=7.0 ACC=20 DEC=20
MOVL C00012 V=7.0 ACC=20 DEC=20
MOVL C00013 V=7.0 ACC=20 DEC=20
MOVL C00014 V=7.0 ACC=20 DEC=20
MOVL C00015 V=7.0 ACC=20 DEC=20
MOVL C00016 V=7.0 ACC=20 DEC=20
MOVL C00017 V=7.0 ACC=20 DEC=20
MOVL C00018 V=7.0 ACC=20 DEC=20
MOVL C00019 V=7.0 ACC=20 DEC=20
MOVL C00020 V=7.0 ACC=20 DEC=20
MOVL C00021 V=7.0 ACC=20 DEC=20
MOVL C00022 V=7.0 ACC=20 DEC=20
MOVC C00023 V=7.0 ACC=20 DEC=20
MOVC C00024 V=7.0 ACC=20 DEC=20
MOVC C00025 V=7.0 ACC=20 DEC=20
MOVL C00026 V=7.0 ACC=20 DEC=20
MOVL C00027 V=7.0 ACC=20 DEC=20
MOVL C00028 V=7.0 ACC=20 DEC=20
MOVL C00029 V=7.0 ACC=20 DEC=20
MOVL C00030 V=7.0 ACC=20 DEC=20
MOVL C00031 V=7.0 ACC=20 DEC=20
MOVL C00032 V=7.0 ACC=20 DEC=20
MOVL C00033 V=7.0 ACC=20 DEC=20
MOVL C00034 V=7.0 ACC=20 DEC=20
MOVL C00035 V=7.0 ACC=20 DEC=20
MOVL C00036 V=7.0 ACC=20 DEC=20
MOVL C00037 V=7.0 ACC=20 DEC=20
MOVL C00038 V=7.0 ACC=20 DEC=20
MOVL C00039 V=7.0 ACC=20 DEC=20
MOVL C00040 V=7.0 ACC=20 DEC=20
MOVL C00041 V=7.0 ACC=20 DEC=20
MOVL C00042 V=7.0 ACC=20 DEC=20
MOVL C00043 V=7.0 ACC=20 DEC=20
MOVL C00044 V=7.0 ACC=20 DEC=20
MOVL C00045 V=7.0 ACC=20 DEC=20
ARCOF
TIMER T=30.00
*LAG2
MOVL C00046 V=11.0 ACC=20 DEC=20
MACRO1 MJ#(0) ARGF2
ARCON
MOVL C00047 V=7.0 ACC=20 DEC=20
MOVL C00048 V=7.0 ACC=20 DEC=20
MOVL C00049 V=7.0 ACC=20 DEC=20
MOVL C00050 V=7.0 ACC=20 DEC=20
MOVL C00051 V=7.0 ACC=20 DEC=20
MOVL C00052 V=7.0 ACC=20 DEC=20
MOVL C00053 V=7.0 ACC=20 DEC=20
MOVL C00054 V=7.0 ACC=20 DEC=20
MOVL C00055 V=7.0 ACC=20 DEC=20
MOVL C00056 V=7.0 ACC=20 DEC=20
MOVL C00057 V=7.0 ACC=20 DEC=20
MOVL C00058 V=7.0 ACC=20 DEC=20
MOVL C00059 V=7.0 ACC=20 DEC=20
MOVL C00060 V=7.0 ACC=20 DEC=20
MOVL C00061 V=7.0 ACC=20 DEC=20
MOVL C00062 V=7.0 ACC=20 DEC=20
MOVL C00063 V=7.0 ACC=20 DEC=20
MOVL C00064 V=7.0 ACC=20 DEC=20
MOVL C00065 V=7.0 ACC=20 DEC=20
MOVC C00066 V=7.0 ACC=20 DEC=20
MOVC C00067 V=7.0 ACC=20 DEC=20
MOVC C00068 V=7.0 ACC=20 DEC=20
MOVL C00069 V=7.0 ACC=20 DEC=20
MOVL C00070 V=7.0 ACC=20 DEC=20
MOVL C00071 V=7.0 ACC=20 DEC=20
MOVL C00072 V=7.0 ACC=20 DEC=20
MOVL C00073 V=7.0 ACC=20 DEC=20
MOVL C00074 V=7.0 ACC=20 DEC=20
MOVL C00075 V=7.0 ACC=20 DEC=20
MOVL C00076 V=7.0 ACC=20 DEC=20
MOVL C00077 V=7.0 ACC=20 DEC=20
MOVL C00078 V=7.0 ACC=20 DEC=20
MOVL C00079 V=7.0 ACC=20 DEC=20
MOVL C00080 V=7.0 ACC=20 DEC=20
MOVL C00081 V=7.0 ACC=20 DEC=20
MOVL C00082 V=7.0 ACC=20 DEC=20
MOVL C00083 V=7.0 ACC=20 DEC=20
MOVL C00084 V=7.0 ACC=20 DEC=20
MOVL C00085 V=7.0 ACC=20 DEC=20
MOVL C00086 V=7.0 ACC=20 DEC=20
MOVL C00087 V=7.0 ACC=20 DEC=20
MOVL C00088 V=7.0 ACC=20 DEC=20
MOVL C00089 V=7.0 ACC=20 DEC=20
ARCOF
TIMER T=30.00
*LAG3
MOVL C00090 V=11.0 ACC=20 DEC=20
MACRO1 MJ#(0) ARGF2
ARCON
MOVL C00091 V=7.0 ACC=20 DEC=20
MOVL C00092 V=7.0 ACC=20 DEC=20
MOVL C00093 V=7.0 ACC=20 DEC=20
MOVL C00094 V=7.0 ACC=20 DEC=20
MOVL C00095 V=7.0 ACC=20 DEC=20
MOVL C00096 V=7.0 ACC=20 DEC=20
MOVL C00097 V=7.0 ACC=20 DEC=20
MOVL C00098 V=7.0 ACC=20 DEC=20
MOVL C00099 V=7.0 ACC=20 DEC=20
MOVL C00100 V=7.0 ACC=20 DEC=20
MOVL C00101 V=7.0 ACC=20 DEC=20
MOVL C00102 V=7.0 ACC=20 DEC=20
MOVL C00103 V=7.0 ACC=20 DEC=20
MOVL C00104 V=7.0 ACC=20 DEC=20
MOVL C00105 V=7.0 ACC=20 DEC=20
MOVL C00106 V=7.0 ACC=20 DEC=20
MOVL C00107 V=7.0 ACC=20 DEC=20
MOVL C00108 V=7.0 ACC=20 DEC=20
MOVL C00109 V=7.0 ACC=20 DEC=20
MOVL C00110 V=7.0 ACC=20 DEC=20
MOVC C00111 V=7.0 ACC=20 DEC=20
MOVC C00112 V=7.0 ACC=20 DEC=20
MOVC C00113 V=7.0 ACC=20 DEC=20
MOVL C00114 V=7.0 ACC=20 DEC=20
MOVL C00115 V=7.0 ACC=20 DEC=20
MOVL C00116 V=7.0 ACC=20 DEC=20
MOVL C00117 V=7.0 ACC=20 DEC=20
MOVL C00118 V=7.0 ACC=20 DEC=20
MOVL C00119 V=7.0 ACC=20 DEC=20
MOVL C00120 V=7.0 ACC=20 DEC=20
MOVL C00121 V=7.0 ACC=20 DEC=20
MOVL C00122 V=7.0 ACC=20 DEC=20
MOVL C00123 V=7.0 ACC=20 DEC=20
MOVL C00124 V=7.0 ACC=20 DEC=20
MOVL C00125 V=7.0 ACC=20 DEC=20
MOVL C00126 V=7.0 ACC=20 DEC=20
MOVL C00127 V=7.0 ACC=20 DEC=20
MOVL C00128 V=7.0 ACC=20 DEC=20
MOVL C00129 V=7.0 ACC=20 DEC=20
MOVL C00130 V=7.0 ACC=20 DEC=20
MOVL C00131 V=7.0 ACC=20 DEC=20
MOVL C00132 V=7.0 ACC=20 DEC=20
MOVL C00133 V=7.0 ACC=20 DEC=20
ARCOF
TIMER T=30.00
*LAG4
MOVL C00134 V=11.0 ACC=20 DEC=20
MACRO1 MJ#(0) ARGF2
ARCON
MOVL C00135 V=7.0 ACC=20 DEC=20
MOVL C00136 V=7.0 ACC=20 DEC=20
MOVL C00137 V=7.0 ACC=20 DEC=20
MOVL C00138 V=7.0 ACC=20 DEC=20
MOVL C00139 V=7.0 ACC=20 DEC=20
MOVL C00140 V=7.0 ACC=20 DEC=20
MOVL C00141 V=7.0 ACC=20 DEC=20
MOVL C00142 V=7.0 ACC=20 DEC=20
MOVL C00143 V=7.0 ACC=20 DEC=20
MOVL C00144 V=7.0 ACC=20 DEC=20
MOVL C00145 V=7.0 ACC=20 DEC=20
MOVL C00146 V=7.0 ACC=20 DEC=20
MOVL C00147 V=7.0 ACC=20 DEC=20
MOVL C00148 V=7.0 ACC=20 DEC=20
MOVL C00149 V=7.0 ACC=20 DEC=20
MOVL C00150 V=7.0 ACC=20 DEC=20
MOVL C00151 V=7.0 ACC=20 DEC=20
MOVL C00152 V=7.0 ACC=20 DEC=20
MOVL C00153 V=7.0 ACC=20 DEC=20
MOVC C00154 V=7.0 ACC=20 DEC=20
MOVC C00155 V=7.0 ACC=20 DEC=20
MOVC C00156 V=7.0 ACC=20 DEC=20
MOVL C00157 V=7.0 ACC=20 DEC=20
MOVL C00158 V=7.0 ACC=20 DEC=20
MOVL C00159 V=7.0 ACC=20 DEC=20
MOVL C00160 V=7.0 ACC=20 DEC=20
MOVL C00161 V=7.0 ACC=20 DEC=20
MOVL C00162 V=7.0 ACC=20 DEC=20
MOVL C00163 V=7.0 ACC=20 DEC=20
MOVL C00164 V=7.0 ACC=20 DEC=20
MOVL C00165 V=7.0 ACC=20 DEC=20
MOVL C00166 V=7.0 ACC=20 DEC=20
MOVL C00167 V=7.0 ACC=20 DEC=20
MOVL C00168 V=7.0 ACC=20 DEC=20
MOVL C00169 V=7.0 ACC=20 DEC=20
MOVL C00170 V=7.0 ACC=20 DEC=20
MOVL C00171 V=7.0 ACC=20 DEC=20
MOVL C00172 V=7.0 ACC=20 DEC=20
MOVL C00173 V=7.0 ACC=20 DEC=20
MOVL C00174 V=7.0 ACC=20 DEC=20
MOVL C00175 V=7.0 ACC=20 DEC=20
MOVL C00176 V=7.0 ACC=20 DEC=20
MOVL C00177 V=7.0 ACC=20 DEC=20
ARCOF
TIMER T=30.00
*LAG5
MOVL C00178 V=11.0 ACC=20 DEC=20
MACRO1 MJ#(0) ARGF2
ARCON
MOVL C00179 V=7.0 ACC=20 DEC=20
MOVL C00180 V=7.0 ACC=20 DEC=20
MOVL C00181 V=7.0 ACC=20 DEC=20
MOVL C00182 V=7.0 ACC=20 DEC=20
MOVL C00183 V=7.0 ACC=20 DEC=20
MOVL C00184 V=7.0 ACC=20 DEC=20
MOVL C00185 V=7.0 ACC=20 DEC=20
MOVL C00186 V=7.0 ACC=20 DEC=20
MOVL C00187 V=7.0 ACC=20 DEC=20
MOVL C00188 V=7.0 ACC=20 DEC=20
MOVL C00189 V=7.0 ACC=20 DEC=20
MOVL C00190 V=7.0 ACC=20 DEC=20
MOVL C00191 V=7.0 ACC=20 DEC=20
MOVL C00192 V=7.0 ACC=20 DEC=20
MOVL C00193 V=7.0 ACC=20 DEC=20
MOVL C00194 V=7.0 ACC=20 DEC=20
MOVL C00195 V=7.0 ACC=20 DEC=20
MOVL C00196 V=7.0 ACC=20 DEC=20
MOVL C00197 V=7.0 ACC=20 DEC=20
MOVL C00198 V=7.0 ACC=20 DEC=20
MOVC C00199 V=7.0 ACC=20 DEC=20
MOVC C00200 V=7.0 ACC=20 DEC=20
MOVC C00201 V=7.0 ACC=20 DEC=20
MOVL C00202 V=7.0 ACC=20 DEC=20
MOVL C00203 V=7.0 ACC=20 DEC=20
MOVL C00204 V=7.0 ACC=20 DEC=20
MOVL C00205 V=7.0 ACC=20 DEC=20
MOVL C00206 V=7.0 ACC=20 DEC=20
MOVL C00207 V=7.0 ACC=20 DEC=20
MOVL C00208 V=7.0 ACC=20 DEC=20
MOVL C00209 V=7.0 ACC=20 DEC=20
MOVL C00210 V=7.0 ACC=20 DEC=20
MOVL C00211 V=7.0 ACC=20 DEC=20
MOVL C00212 V=7.0 ACC=20 DEC=20
MOVL C00213 V=7.0 ACC=20 DEC=20
MOVL C00214 V=7.0 ACC=20 DEC=20
MOVL C00215 V=7.0 ACC=20 DEC=20
MOVL C00216 V=7.0 ACC=20 DEC=20
MOVL C00217 V=7.0 ACC=20 DEC=20
MOVL C00218 V=7.0 ACC=20 DEC=20
MOVL C00219 V=7.0 ACC=20 DEC=20
MOVL C00220 V=7.0 ACC=20 DEC=20
MOVL C00221 V=7.0 ACC=20 DEC=20
ARCOF
TIMER T=30.00
*LAG6
MOVL C00222 V=11.0 ACC=20 DEC=20
MACRO1 MJ#(0) ARGF2
ARCON
MOVL C00223 V=7.0 ACC=20 DEC=20
MOVL C00224 V=7.0 ACC=20 DEC=20
MOVL C00225 V=7.0 ACC=20 DEC=20
MOVL C00226 V=7.0 ACC=20 DEC=20
MOVL C00227 V=7.0 ACC=20 DEC=20
MOVL C00228 V=7.0 ACC=20 DEC=20
MOVL C00229 V=7.0 ACC=20 DEC=20
MOVL C00230 V=7.0 ACC=20 DEC=20
MOVL C00231 V=7.0 ACC=20 DEC=20
MOVL C00232 V=7.0 ACC=20 DEC=20
MOVL C00233 V=7.0 ACC=20 DEC=20
MOVL C00234 V=7.0 ACC=20 DEC=20
MOVL C00235 V=7.0 ACC=20 DEC=20
MOVL C00236 V=7.0 ACC=20 DEC=20
MOVL C00237 V=7.0 ACC=20 DEC=20
MOVL C00238 V=7.0 ACC=20 DEC=20
MOVL C00239 V=7.0 ACC=20 DEC=20
MOVL C00240 V=7.0 ACC=20 DEC=20
MOVL C00241 V=7.0 ACC=20 DEC=20
MOVC C00242 V=7.0 ACC=20 DEC=20
MOVC C00243 V=7.0 ACC=20 DEC=20
MOVC C00244 V=7.0 ACC=20 DEC=20
MOVL C00245 V=7.0 ACC=20 DEC=20
MOVL C00246 V=7.0 ACC=20 DEC=20
MOVL C00247 V=7.0 ACC=20 DEC=20
MOVL C00248 V=7.0 ACC=20 DEC=20
MOVL C00249 V=7.0 ACC=20 DEC=20
MOVL C00250 V=7.0 ACC=20 DEC=20
MOVL C00251 V=7.0 ACC=20 DEC=20
MOVL C00252 V=7.0 ACC=20 DEC=20
MOVL C00253 V=7.0 ACC=20 DEC=20
MOVL C00254 V=7.0 ACC=20 DEC=20
MOVL C00255 V=7.0 ACC=20 DEC=20
MOVL C00256 V=7.0 ACC=20 DEC=20
MOVL C00257 V=7.0 ACC=20 DEC=20
MOVL C00258 V=7.0 ACC=20 DEC=20
MOVL C00259 V=7.0 ACC=20 DEC=20
MOVL C00260 V=7.0 ACC=20 DEC=20
MOVL C00261 V=7.0 ACC=20 DEC=20
MOVL C00262 V=7.0 ACC=20 DEC=20
MOVL C00263 V=7.0 ACC=20 DEC=20
MOVL C00264 V=7.0 ACC=20 DEC=20
MOVL C00265 V=7.0 ACC=20 DEC=20
ARCOF
TIMER T=30.00
*LAG7
MOVL C00266 V=11.0 ACC=20 DEC=20
MACRO1 MJ#(0) ARGF2
ARCON
MOVL C00267 V=7.0 ACC=20 DEC=20
MOVL C00268 V=7.0 ACC=20 DEC=20
MOVL C00269 V=7.0 ACC=20 DEC=20
MOVL C00270 V=7.0 ACC=20 DEC=20
MOVL C00271 V=7.0 ACC=20 DEC=20
MOVL C00272 V=7.0 ACC=20 DEC=20
MOVL C00273 V=7.0 ACC=20 DEC=20
MOVL C00274 V=7.0 ACC=20 DEC=20
MOVL C00275 V=7.0 ACC=20 DEC=20
MOVL C00276 V=7.0 ACC=20 DEC=20
MOVL C00277 V=7.0 ACC=20 DEC=20
MOVL C00278 V=7.0 ACC=20 DEC=20
MOVL C00279 V=7.0 ACC=20 DEC=20
MOVL C00280 V=7.0 ACC=20 DEC=20
MOVL C00281 V=7.0 ACC=20 DEC=20
MOVL C00282 V=7.0 ACC=20 DEC=20
MOVL C00283 V=7.0 ACC=20 DEC=20
MOVL C00284 V=7.0 ACC=20 DEC=20
MOVL C00285 V=7.0 ACC=20 DEC=20
MOVL C00286 V=7.0 ACC=20 DEC=20
MOVC C00287 V=7.0 ACC=20 DEC=20
MOVC C00288 V=7.0 ACC=20 DEC=20
MOVC C00289 V=7.0 ACC=20 DEC=20
MOVL C00290 V=7.0 ACC=20 DEC=20
MOVL C00291 V=7.0 ACC=20 DEC=20
MOVL C00292 V=7.0 ACC=20 DEC=20
MOVL C00293 V=7.0 ACC=20 DEC=20
MOVL C00294 V=7.0 ACC=20 DEC=20
MOVL C00295 V=7.0 ACC=20 DEC=20
MOVL C00296 V=7.0 ACC=20 DEC=20
MOVL C00297 V=7.0 ACC=20 DEC=20
MOVL C00298 V=7.0 ACC=20 DEC=20
MOVL C00299 V=7.0 ACC=20 DEC=20
MOVL C00300 V=7.0 ACC=20 DEC=20
MOVL C00301 V=7.0 ACC=20 DEC=20
MOVL C00302 V=7.0 ACC=20 DEC=20
MOVL C00303 V=7.0 ACC=20 DEC=20
MOVL C00304 V=7.0 ACC=20 DEC=20
MOVL C00305 V=7.0 ACC=20 DEC=20
MOVL C00306 V=7.0 ACC=20 DEC=20
MOVL C00307 V=7.0 ACC=20 DEC=20
MOVL C00308 V=7.0 ACC=20 DEC=20
MOVL C00309 V=7.0 ACC=20 DEC=20
ARCOF
TIMER T=30.00
*LAG8
MOVL C00310 V=11.0 ACC=20 DEC=20
MACRO1 MJ#(0) ARGF2
ARCON
MOVL C00311 V=7.0 ACC=20 DEC=20
MOVL C00312 V=7.0 ACC=20 DEC=20
MOVL C00313 V=7.0 ACC=20 DEC=20
MOVL C00314 V=7.0 ACC=20 DEC=20
MOVL C00315 V=7.0 ACC=20 DEC=20
MOVL C00316 V=7.0 ACC=20 DEC=20
MOVL C00317 V=7.0 ACC=20 DEC=20
MOVL C00318 V=7.0 ACC=20 DEC=20
MOVL C00319 V=7.0 ACC=20 DEC=20
MOVL C00320 V=7.0 ACC=20 DEC=20
MOVL C00321 V=7.0 ACC=20 DEC=20
MOVL C00322 V=7.0 ACC=20 DEC=20
MOVL C00323 V=7.0 ACC=20 DEC=20
MOVL C00324 V=7.0 ACC=20 DEC=20
MOVL C00325 V=7.0 ACC=20 DEC=20
MOVL C00326 V=7.0 ACC=20 DEC=20
MOVL C00327 V=7.0 ACC=20 DEC=20
MOVL C00328 V=7.0 ACC=20 DEC=20
MOVL C00329 V=7.0 ACC=20 DEC=20
MOVC C00330 V=7.0 ACC=20 DEC=20
MOVC C00331 V=7.0 ACC=20 DEC=20
MOVC C00332 V=7.0 ACC=20 DEC=20
MOVL C00333 V=7.0 ACC=20 DEC=20
MOVL C00334 V=7.0 ACC=20 DEC=20
MOVL C00335 V=7.0 ACC=20 DEC=20
MOVL C00336 V=7.0 ACC=20 DEC=20
MOVL C00337 V=7.0 ACC=20 DEC=20
MOVL C00338 V=7.0 ACC=20 DEC=20
MOVL C00339 V=7.0 ACC=20 DEC=20
MOVL C00340 V=7.0 ACC=20 DEC=20
MOVL C00341 V=7.0 ACC=20 DEC=20
MOVL C00342 V=7.0 ACC=20 DEC=20
MOVL C00343 V=7.0 ACC=20 DEC=20
MOVL C00344 V=7.0 ACC=20 DEC=20
MOVL C00345 V=7.0 ACC=20 DEC=20
MOVL C00346 V=7.0 ACC=20 DEC=20
MOVL C00347 V=7.0 ACC=20 DEC=20
MOVL C00348 V=7.0 ACC=20 DEC=20
MOVL C00349 V=7.0 ACC=20 DEC=20
MOVL C00350 V=7.0 ACC=20 DEC=20
MOVL C00351 V=7.0 ACC=20 DEC=20
MOVL C00352 V=7.0 ACC=20 DEC=20
MOVL C00353 V=7.0 ACC=20 DEC=20
ARCOF
TIMER T=30.00
*LAG9
MOVL C00354 V=11.0 ACC=20 DEC=20
MACRO1 MJ#(0) ARGF2
ARCON
MOVL C00355 V=7.0 ACC=20 DEC=20
MOVL C00356 V=7.0 ACC=20 DEC=20
MOVL C00357 V=7.0 ACC=20 DEC=20
MOVL C00358 V=7.0 ACC=20 DEC=20
MOVL C00359 V=7.0 ACC=20 DEC=20
MOVL C00360 V=7.0 ACC=20 DEC=20
MOVL C00361 V=7.0 ACC=20 DEC=20
MOVL C00362 V=7.0 ACC=20 DEC=20
MOVL C00363 V=7.0 ACC=20 DEC=20
MOVL C00364 V=7.0 ACC=20 DEC=20
MOVL C00365 V=7.0 ACC=20 DEC=20
MOVL C00366 V=7.0 ACC=20 DEC=20
MOVL C00367 V=7.0 ACC=20 DEC=20
MOVL C00368 V=7.0 ACC=20 DEC=20
MOVL C00369 V=7.0 ACC=20 DEC=20
MOVL C00370 V=7.0 ACC=20 DEC=20
MOVL C00371 V=7.0 ACC=20 DEC=20
MOVL C00372 V=7.0 ACC=20 DEC=20
MOVL C00373 V=7.0 ACC=20 DEC=20
MOVL C00374 V=7.0 ACC=20 DEC=20
MOVC C00375 V=7.0 ACC=20 DEC=20
MOVC C00376 V=7.0 ACC=20 DEC=20
MOVC C00377 V=7.0 ACC=20 DEC=20
MOVL C00378 V=7.0 ACC=20 DEC=20
MOVL C00379 V=7.0 ACC=20 DEC=20
MOVL C00380 V=7.0 ACC=20 DEC=20
MOVL C00381 V=7.0 ACC=20 DEC=20
MOVL C00382 V=7.0 ACC=20 DEC=20
MOVL C00383 V=7.0 ACC=20 DEC=20
MOVL C00384 V=7.0 ACC=20 DEC=20
MOVL C00385 V=7.0 ACC=20 DEC=20
MOVL C00386 V=7.0 ACC=20 DEC=20
MOVL C00387 V=7.0 ACC=20 DEC=20
MOVL C00388 V=7.0 ACC=20 DEC=20
MOVL C00389 V=7.0 ACC=20 DEC=20
MOVL C00390 V=7.0 ACC=20 DEC=20
MOVL C00391 V=7.0 ACC=20 DEC=20
MOVL C00392 V=7.0 ACC=20 DEC=20
MOVL C00393 V=7.0 ACC=20 DEC=20
MOVL C00394 V=7.0 ACC=20 DEC=20
MOVL C00395 V=7.0 ACC=20 DEC=20
MOVL C00396 V=7.0 ACC=20 DEC=20
MOVL C00397 V=7.0 ACC=20 DEC=20
ARCOF
TIMER T=30.00
*LAG10
MOVL C00398 V=11.0 ACC=20 DEC=20
MACRO1 MJ#(0) ARGF2
ARCON
MOVL C00399 V=7.0 ACC=20 DEC=20
MOVL C00400 V=7.0 ACC=20 DEC=20
MOVL C00401 V=7.0 ACC=20 DEC=20
MOVL C00402 V=7.0 ACC=20 DEC=20
MOVL C00403 V=7.0 ACC=20 DEC=20
MOVL C00404 V=7.0 ACC=20 DEC=20
MOVL C00405 V=7.0 ACC=20 DEC=20
MOVL C00406 V=7.0 ACC=20 DEC=20
MOVL C00407 V=7.0 ACC=20 DEC=20
MOVL C00408 V=7.0 ACC=20 DEC=20
MOVL C00409 V=7.0 ACC=20 DEC=20
MOVL C00410 V=7.0 ACC=20 DEC=20
MOVL C00411 V=7.0 ACC=20 DEC=20
MOVL C00412 V=7.0 ACC=20 DEC=20
MOVL C00413 V=7.0 ACC=20 DEC=20
MOVL C00414 V=7.0 ACC=20 DEC=20
MOVL C00415 V=7.0 ACC=20 DEC=20
MOVL C00416 V=7.0 ACC=20 DEC=20
MOVL C00417 V=7.0 ACC=20 DEC=20
MOVC C00418 V=7.0 ACC=20 DEC=20
MOVC C00419 V=7.0 ACC=20 DEC=20
MOVC C00420 V=7.0 ACC=20 DEC=20
MOVL C00421 V=7.0 ACC=20 DEC=20
MOVL C00422 V=7.0 ACC=20 DEC=20
MOVL C00423 V=7.0 ACC=20 DEC=20
MOVL C00424 V=7.0 ACC=20 DEC=20
MOVL C00425 V=7.0 ACC=20 DEC=20
MOVL C00426 V=7.0 ACC=20 DEC=20
MOVL C00427 V=7.0 ACC=20 DEC=20
MOVL C00428 V=7.0 ACC=20 DEC=20
MOVL C00429 V=7.0 ACC=20 DEC=20
MOVL C00430 V=7.0 ACC=20 DEC=20
MOVL C00431 V=7.0 ACC=20 DEC=20
MOVL C00432 V=7.0 ACC=20 DEC=20
MOVL C00433 V=7.0 ACC=20 DEC=20
MOVL C00434 V=7.0 ACC=20 DEC=20
MOVL C00435 V=7.0 ACC=20 DEC=20
MOVL C00436 V=7.0 ACC=20 DEC=20
MOVL C00437 V=7.0 ACC=20 DEC=20
MOVL C00438 V=7.0 ACC=20 DEC=20
MOVL C00439 V=7.0 ACC=20 DEC=20
MOVL C00440 V=7.0 ACC=20 DEC=20
MOVL C00441 V=7.0 ACC=20 DEC=20
ARCOF
TIMER T=30.00
*LAG11
MOVL C00442 V=11.0 ACC=20 DEC=20
MACRO1 MJ#(0) ARGF2
ARCON
MOVL C00443 V=7.0 ACC=20 DEC=20
MOVL C00444 V=7.0 ACC=20 DEC=20
MOVL C00445 V=7.0 ACC=20 DEC=20
MOVL C00446 V=7.0 ACC=20 DEC=20
MOVL C00447 V=7.0 ACC=20 DEC=20
MOVL C00448 V=7.0 ACC=20 DEC=20
MOVL C00449 V=7.0 ACC=20 DEC=20
MOVL C00450 V=7.0 ACC=20 DEC=20
MOVL C00451 V=7.0 ACC=20 DEC=20
MOVL C00452 V=7.0 ACC=20 DEC=20
MOVL C00453 V=7.0 ACC=20 DEC=20
MOVL C00454 V=7.0 ACC=20 DEC=20
MOVL C00455 V=7.0 ACC=20 DEC=20
MOVL C00456 V=7.0 ACC=20 DEC=20
MOVL C00457 V=7.0 ACC=20 DEC=20
MOVL C00458 V=7.0 ACC=20 DEC=20
MOVL C00459 V=7.0 ACC=20 DEC=20
MOVL C00460 V=7.0 ACC=20 DEC=20
MOVL C00461 V=7.0 ACC=20 DEC=20
MOVL C00462 V=7.0 ACC=20 DEC=20
MOVC C00463 V=7.0 ACC=20 DEC=20
MOVC C00464 V=7.0 ACC=20 DEC=20
MOVC C00465 V=7.0 ACC=20 DEC=20
MOVL C00466 V=7.0 ACC=20 DEC=20
MOVL C00467 V=7.0 ACC=20 DEC=20
MOVL C00468 V=7.0 ACC=20 DEC=20
MOVL C00469 V=7.0 ACC=20 DEC=20
MOVL C00470 V=7.0 ACC=20 DEC=20
MOVL C00471 V=7.0 ACC=20 DEC=20
MOVL C00472 V=7.0 ACC=20 DEC=20
MOVL C00473 V=7.0 ACC=20 DEC=20
MOVL C00474 V=7.0 ACC=20 DEC=20
MOVL C00475 V=7.0 ACC=20 DEC=20
MOVL C00476 V=7.0 ACC=20 DEC=20
MOVL C00477 V=7.0 ACC=20 DEC=20
MOVL C00478 V=7.0 ACC=20 DEC=20
MOVL C00479 V=7.0 ACC=20 DEC=20
MOVL C00480 V=7.0 ACC=20 DEC=20
MOVL C00481 V=7.0 ACC=20 DEC=20
MOVL C00482 V=7.0 ACC=20 DEC=20
MOVL C00483 V=7.0 ACC=20 DEC=20
MOVL C00484 V=7.0 ACC=20 DEC=20
MOVL C00485 V=7.0 ACC=20 DEC=20
ARCOF
TIMER T=30.00
*LAG12
MOVL C00486 V=11.0 ACC=20 DEC=20
MACRO1 MJ#(0) ARGF2
ARCON
MOVL C00487 V=7.0 ACC=20 DEC=20
MOVL C00488 V=7.0 ACC=20 DEC=20
MOVL C00489 V=7.0 ACC=20 DEC=20
MOVL C00490 V=7.0 ACC=20 DEC=20
MOVL C00491 V=7.0 ACC=20 DEC=20
MOVL C00492 V=7.0 ACC=20 DEC=20
MOVL C00493 V=7.0 ACC=20 DEC=20
MOVL C00494 V=7.0 ACC=20 DEC=20
MOVL C00495 V=7.0 ACC=20 DEC=20
MOVL C00496 V=7.0 ACC=20 DEC=20
MOVL C00497 V=7.0 ACC=20 DEC=20
MOVL C00498 V=7.0 ACC=20 DEC=20
MOVL C00499 V=7.0 ACC=20 DEC=20
MOVL C00500 V=7.0 ACC=20 DEC=20
MOVL C00501 V=7.0 ACC=20 DEC=20
MOVL C00502 V=7.0 ACC=20 DEC=20
MOVL C00503 V=7.0 ACC=20 DEC=20
MOVL C00504 V=7.0 ACC=20 DEC=20
MOVL C00505 V=7.0 ACC=20 DEC=20
MOVC C00506 V=7.0 ACC=20 DEC=20
MOVC C00507 V=7.0 ACC=20 DEC=20
MOVC C00508 V=7.0 ACC=20 DEC=20
MOVL C00509 V=7.0 ACC=20 DEC=20
MOVL C00510 V=7.0 ACC=20 DEC=20
MOVL C00511 V=7.0 ACC=20 DEC=20
MOVL C00512 V=7.0 ACC=20 DEC=20
MOVL C00513 V=7.0 ACC=20 DEC=20
MOVL C00514 V=7.0 ACC=20 DEC=20
MOVL C00515 V=7.0 ACC=20 DEC=20
MOVL C00516 V=7.0 ACC=20 DEC=20
MOVL C00517 V=7.0 ACC=20 DEC=20
MOVL C00518 V=7.0 ACC=20 DEC=20
MOVL C00519 V=7.0 ACC=20 DEC=20
MOVL C00520 V=7.0 ACC=20 DEC=20
MOVL C00521 V=7.0 ACC=20 DEC=20
MOVL C00522 V=7.0 ACC=20 DEC=20
MOVL C00523 V=7.0 ACC=20 DEC=20
MOVL C00524 V=7.0 ACC=20 DEC=20
MOVL C00525 V=7.0 ACC=20 DEC=20
MOVL C00526 V=7.0 ACC=20 DEC=20
MOVL C00527 V=7.0 ACC=20 DEC=20
MOVL C00528 V=7.0 ACC=20 DEC=20
MOVL C00529 V=7.0 ACC=20 DEC=20
ARCOF
TIMER T=30.00
*LAG13
MOVL C00530 V=11.0 ACC=20 DEC=20
MACRO1 MJ#(0) ARGF2
ARCON
MOVL C00531 V=7.0 ACC=20 DEC=20
MOVL C00532 V=7.0 ACC=20 DEC=20
MOVL C00533 V=7.0 ACC=20 DEC=20
MOVL C00534 V=7.0 ACC=20 DEC=20
MOVL C00535 V=7.0 ACC=20 DEC=20
MOVL C00536 V=7.0 ACC=20 DEC=20
MOVL C00537 V=7.0 ACC=20 DEC=20
MOVL C00538 V=7.0 ACC=20 DEC=20
MOVL C00539 V=7.0 ACC=20 DEC=20
MOVL C00540 V=7.0 ACC=20 DEC=20
MOVL C00541 V=7.0 ACC=20 DEC=20
MOVL C00542 V=7.0 ACC=20 DEC=20
MOVL C00543 V=7.0 ACC=20 DEC=20
MOVL C00544 V=7.0 ACC=20 DEC=20
MOVL C00545 V=7.0 ACC=20 DEC=20
MOVL C00546 V=7.0 ACC=20 DEC=20
MOVL C00547 V=7.0 ACC=20 DEC=20
MOVL C00548 V=7.0 ACC=20 DEC=20
MOVL C00549 V=7.0 ACC=20 DEC=20
MOVL C00550 V=7.0 ACC=20 DEC=20
MOVC C00551 V=7.0 ACC=20 DEC=20
MOVC C00552 V=7.0 ACC=20 DEC=20
MOVC C00553 V=7.0 ACC=20 DEC=20
MOVL C00554 V=7.0 ACC=20 DEC=20
MOVL C00555 V=7.0 ACC=20 DEC=20
MOVL C00556 V=7.0 ACC=20 DEC=20
MOVL C00557 V=7.0 ACC=20 DEC=20
MOVL C00558 V=7.0 ACC=20 DEC=20
MOVL C00559 V=7.0 ACC=20 DEC=20
MOVL C00560 V=7.0 ACC=20 DEC=20
MOVL C00561 V=7.0 ACC=20 DEC=20
MOVL C00562 V=7.0 ACC=20 DEC=20
MOVL C00563 V=7.0 ACC=20 DEC=20
MOVL C00564 V=7.0 ACC=20 DEC=20
MOVL C00565 V=7.0 ACC=20 DEC=20
MOVL C00566 V=7.0 ACC=20 DEC=20
MOVL C00567 V=7.0 ACC=20 DEC=20
MOVL C00568 V=7.0 ACC=20 DEC=20
MOVL C00569 V=7.0 ACC=20 DEC=20
MOVL C00570 V=7.0 ACC=20 DEC=20
MOVL C00571 V=7.0 ACC=20 DEC=20
MOVL C00572 V=7.0 ACC=20 DEC=20
MOVL C00573 V=7.0 ACC=20 DEC=20
ARCOF
TIMER T=30.00
*LAG14
MOVL C00574 V=11.0 ACC=20 DEC=20
MACRO1 MJ#(0) ARGF2
ARCON
MOVL C00575 V=7.0 ACC=20 DEC=20
MOVL C00576 V=7.0 ACC=20 DEC=20
MOVL C00577 V=7.0 ACC=20 DEC=20
MOVL C00578 V=7.0 ACC=20 DEC=20
MOVL C00579 V=7.0 ACC=20 DEC=20
MOVL C00580 V=7.0 ACC=20 DEC=20
MOVL C00581 V=7.0 ACC=20 DEC=20
MOVL C00582 V=7.0 ACC=20 DEC=20
MOVL C00583 V=7.0 ACC=20 DEC=20
MOVL C00584 V=7.0 ACC=20 DEC=20
MOVL C00585 V=7.0 ACC=20 DEC=20
MOVL C00586 V=7.0 ACC=20 DEC=20
MOVL C00587 V=7.0 ACC=20 DEC=20
MOVL C00588 V=7.0 ACC=20 DEC=20
MOVL C00589 V=7.0 ACC=20 DEC=20
MOVL C00590 V=7.0 ACC=20 DEC=20
MOVL C00591 V=7.0 ACC=20 DEC=20
MOVL C00592 V=7.0 ACC=20 DEC=20
MOVL C00593 V=7.0 ACC=20 DEC=20
MOVC C00594 V=7.0 ACC=20 DEC=20
MOVC C00595 V=7.0 ACC=20 DEC=20
MOVC C00596 V=7.0 ACC=20 DEC=20
MOVL C00597 V=7.0 ACC=20 DEC=20
MOVL C00598 V=7.0 ACC=20 DEC=20
MOVL C00599 V=7.0 ACC=20 DEC=20
MOVL C00600 V=7.0 ACC=20 DEC=20
MOVL C00601 V=7.0 ACC=20 DEC=20
MOVL C00602 V=7.0 ACC=20 DEC=20
MOVL C00603 V=7.0 ACC=20 DEC=20
MOVL C00604 V=7.0 ACC=20 DEC=20
MOVL C00605 V=7.0 ACC=20 DEC=20
MOVL C00606 V=7.0 ACC=20 DEC=20
MOVL C00607 V=7.0 ACC=20 DEC=20
MOVL C00608 V=7.0 ACC=20 DEC=20
MOVL C00609 V=7.0 ACC=20 DEC=20
MOVL C00610 V=7.0 ACC=20 DEC=20
MOVL C00611 V=7.0 ACC=20 DEC=20
MOVL C00612 V=7.0 ACC=20 DEC=20
MOVL C00613 V=7.0 ACC=20 DEC=20
MOVL C00614 V=7.0 ACC=20 DEC=20
MOVL C00615 V=7.0 ACC=20 DEC=20
MOVL C00616 V=7.0 ACC=20 DEC=20
MOVL C00617 V=7.0 ACC=20 DEC=20
ARCOF
TIMER T=30.00
*LAG15
MOVL C00618 V=11.0 ACC=20 DEC=20
MACRO1 MJ#(0) ARGF2
ARCON
MOVL C00619 V=7.0 ACC=20 DEC=20
MOVL C00620 V=7.0 ACC=20 DEC=20
MOVL C00621 V=7.0 ACC=20 DEC=20
MOVL C00622 V=7.0 ACC=20 DEC=20
MOVL C00623 V=7.0 ACC=20 DEC=20
MOVL C00624 V=7.0 ACC=20 DEC=20
MOVL C00625 V=7.0 ACC=20 DEC=20
MOVL C00626 V=7.0 ACC=20 DEC=20
MOVL C00627 V=7.0 ACC=20 DEC=20
MOVL C00628 V=7.0 ACC=20 DEC=20
MOVL C00629 V=7.0 ACC=20 DEC=20
MOVL C00630 V=7.0 ACC=20 DEC=20
MOVL C00631 V=7.0 ACC=20 DEC=20
MOVL C00632 V=7.0 ACC=20 DEC=20
MOVL C00633 V=7.0 ACC=20 DEC=20
MOVL C00634 V=7.0 ACC=20 DEC=20
MOVL C00635 V=7.0 ACC=20 DEC=20
MOVL C00636 V=7.0 ACC=20 DEC=20
MOVL C00637 V=7.0 ACC=20 DEC=20
MOVL C00638 V=7.0 ACC=20 DEC=20
MOVC C00639 V=7.0 ACC=20 DEC=20
MOVC C00640 V=7.0 ACC=20 DEC=20
MOVC C00641 V=7.0 ACC=20 DEC=20
MOVL C00642 V=7.0 ACC=20 DEC=20
MOVL C00643 V=7.0 ACC=20 DEC=20
MOVL C00644 V=7.0 ACC=20 DEC=20
MOVL C00645 V=7.0 ACC=20 DEC=20
MOVL C00646 V=7.0 ACC=20 DEC=20
MOVL C00647 V=7.0 ACC=20 DEC=20
MOVL C00648 V=7.0 ACC=20 DEC=20
MOVL C00649 V=7.0 ACC=20 DEC=20
MOVL C00650 V=7.0 ACC=20 DEC=20
MOVL C00651 V=7.0 ACC=20 DEC=20
MOVL C00652 V=7.0 ACC=20 DEC=20
MOVL C00653 V=7.0 ACC=20 DEC=20
MOVL C00654 V=7.0 ACC=20 DEC=20
MOVL C00655 V=7.0 ACC=20 DEC=20
MOVL C00656 V=7.0 ACC=20 DEC=20
MOVL C00657 V=7.0 ACC=20 DEC=20
MOVL C00658 V=7.0 ACC=20 DEC=20
MOVL C00659 V=7.0 ACC=20 DEC=20
MOVL C00660 V=7.0 ACC=20 DEC=20
MOVL C00661 V=7.0 ACC=20 DEC=20
ARCOF
TIMER T=30.00
MOVL C00662 V=11.0 ACC=20 DEC=20
MOVJ C00663 VJ=0.78
END
